(* IEC 61131-3 sources: plc-vscode/tests/st/test-ready/trust-platform/examples/communication/multi_driver/src, 2 files *)

(* ---- config.st ---- *)
CONFIGURATION Config
RESOURCE CommRes ON PLC
    TASK MainTask (INTERVAL := T#100ms, PRIORITY := 1);
    PROGRAM P1 WITH MainTask : Main;
END_RESOURCE
VAR_CONFIG
    P1.DI0 AT %IX0.0 : BOOL;
    P1.DO0 AT %QX0.0 : BOOL;
END_VAR
END_CONFIGURATION

(* ---- main.st ---- *)
PROGRAM Main
VAR
    DI0 : BOOL;
    DO0 : BOOL;
END_VAR

DO0 := DI0;
END_PROGRAM
